// TIA Portal V21 export
// export: Created 2026-11-11T00:47:54.924807Z, ExportSetting WithDefaults, DisplayName Totally Integrated Automation Portal, DisplayVersion V21 Update 3, DisplayName STEP 7 Professional, DisplayVersion V21 Update 3, DisplayName STEP 7 Safety, DisplayVersion V21, DisplayName Tech WebApplication, DisplayVersion V21, DisplayName WinCC Basic/Comfort/Advanced, DisplayVersion V21 Update 3, DisplayName WinCC Unified, DisplayVersion V21 Update 3
FUNCTION_BLOCK "FB_Lad_ou005"   // FB346, LAD
{ S7_Optimized_Access := 'TRUE' }
VERSION : 0.1
// stored: AutoNumber true, IsIECCheckEnabled false, IsRetainMemResEnabled false, MemoryReserve 100, SetENOAutomatically false, UDAEnableTagReadback false
   VAR_INPUT
      v_req : Bool;
      v_to_s : String;
      v_cc : String;
      v_subject : String;
      v_text : String;
      v_attachment : Array[0..99] of Byte;
      v_attachment_name : String;
      v_mail_addr_param : Array[0..99] of Byte;
   END_VAR
   VAR_OUTPUT
      v_done : Bool;
      v_busy : Bool;
      v_error : Bool;
      v_status : Word;
   END_VAR
   VAR
      inst { S7_SetPoint := 'True'} : TMAIL_C;
   END_VAR
BEGIN

REGION Network 1: Description of TMAIL_C
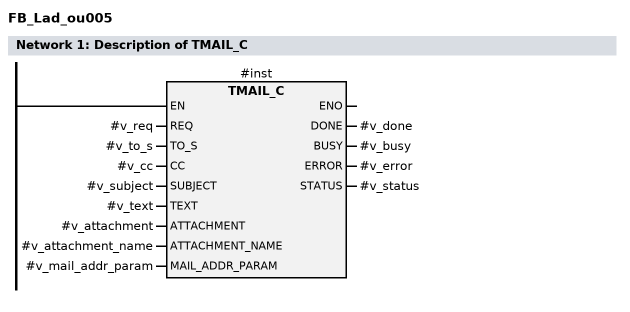
   RUNG wire#powerrail
      #inst.TMAIL_C(REQ := #v_req, TO_S := #v_to_s, CC := #v_cc, SUBJECT := #v_subject, TEXT := #v_text, ATTACHMENT := #v_attachment, ATTACHMENT_NAME := #v_attachment_name, MAIL_ADDR_PARAM := #v_mail_addr_param, DONE => #v_done, BUSY => #v_busy, ERROR => #v_error, STATUS => #v_status)
   END_RUNG
   // the same network as SCL:
   #inst(REQ := #v_req,   // TMAIL_C
         TO_S := #v_to_s,
         CC := #v_cc,
         SUBJECT := #v_subject,
         TEXT := #v_text,
         ATTACHMENT := #v_attachment,
         ATTACHMENT_NAME := #v_attachment_name,
         MAIL_ADDR_PARAM := #v_mail_addr_param,
         DONE => #v_done,
         BUSY => #v_busy,
         ERROR => #v_error,
         STATUS => #v_status);
END_REGION
END_FUNCTION_BLOCK
